// TIA Portal V21 export
// export: Created 2026-11-03T19:44:49.0635428Z, ExportSetting WithDefaults, WithReadOnly, DisplayName Totally Integrated Automation Portal, DisplayVersion V21, DisplayName STEP 7 Professional, DisplayVersion V21, DisplayName STEP 7 Safety, DisplayVersion V21, DisplayName Tech WebApplication, DisplayVersion V21, DisplayName WinCC Basic/Comfort/Advanced, DisplayVersion V21, DisplayName WinCC Professional, DisplayVersion V21, DisplayName WinCC Unified, DisplayVersion V21
DATA_BLOCK "DB_FAT_Demo"   // DB1
{ S7_Optimized_Access := 'FALSE' }
VERSION : 1.0
// SPDX-License-Identifier: MIT. Public passive laboratory example.
// stored: AutoNumber true, CodeModifiedDate 2026-11-03T19:44:32.7091278Z, CompileDate 2026-11-03T19:44:33.4739621Z, CreationDate 2026-11-03T19:44:31.2051572Z, DBAccessibleFromOPCUA true, DBAccessibleFromWebserver true, DownloadDate 0001-01-01T00:00:00Z, InterfaceModifiedDate 2026-11-03T19:44:32.7091278Z, IsConsistent true, IsKnowHowProtected false, IsOnlyStoredInLoadMemory false, IsPLCDB false, IsWriteProtectedInAS false, LoadMemoryLength 5286, ModifiedDate 2026-11-03T19:44:32.7091278Z, ParameterModified 2026-11-03T19:44:32.7091278Z, StructureModified 2026-11-03T19:44:32.7091278Z, WorkMemoryLength 192
   VAR RETAIN
      EnableDemo { ExternalAccessible := 'False'; ExternalVisible := 'False'; ExternalWritable := 'False'} : Bool := TRUE;   // isolated virtual copy only
      StopHealthy : Bool := TRUE;
      P101_Request : Bool := FALSE;
      P101_RequestedSpeed : Real := REAL#60.0;
      P101_RunCommand { ExternalWritable := 'False'} : Bool := FALSE;
      P101_SpeedCommand { ExternalWritable := 'False'} : Real := REAL#0.0;
      P101_Running : Bool := FALSE;
      P101_SpeedFeedback : Real := REAL#0.0;
      P101_Fault : Bool := FALSE;
      P201_Request : Bool := FALSE;
      P201_RequestedSpeed : Real := REAL#60.0;
      P201_RunCommand { ExternalWritable := 'False'} : Bool := FALSE;
      P201_SpeedCommand { ExternalWritable := 'False'} : Real := REAL#0.0;
      P201_Running : Bool := FALSE;
      P201_SpeedFeedback : Real := REAL#0.0;
      P201_Fault : Bool := FALSE;
      P202_Request : Bool := FALSE;
      P202_RequestedSpeed : Real := REAL#60.0;
      P202_RunCommand { ExternalWritable := 'False'} : Bool := FALSE;
      P202_SpeedCommand { ExternalWritable := 'False'} : Real := REAL#0.0;
      P202_Running : Bool := FALSE;
      P202_SpeedFeedback : Real := REAL#0.0;
      P202_Fault : Bool := FALSE;
      P301_Request : Bool := FALSE;
      P301_RequestedSpeed : Real := REAL#60.0;
      P301_RunCommand { ExternalWritable := 'False'} : Bool := FALSE;
      P301_SpeedCommand { ExternalWritable := 'False'} : Real := REAL#0.0;
      P301_Running : Bool := FALSE;
      P301_SpeedFeedback : Real := REAL#0.0;
      P301_Fault : Bool := FALSE;
      XV101_Request : Bool := FALSE;
      XV101_OpenCommand { ExternalWritable := 'False'} : Bool := FALSE;
      XV101_Open : Bool := FALSE;
      XV101_Closed : Bool := TRUE;
      XV201_Request : Bool := FALSE;
      XV201_OpenCommand { ExternalWritable := 'False'} : Bool := FALSE;
      XV201_Open : Bool := FALSE;
      XV201_Closed : Bool := TRUE;
      XV202_Request : Bool := FALSE;
      XV202_OpenCommand { ExternalWritable := 'False'} : Bool := FALSE;
      XV202_Open : Bool := FALSE;
      XV202_Closed : Bool := TRUE;
      XV301_Request : Bool := FALSE;
      XV301_OpenCommand { ExternalWritable := 'False'} : Bool := FALSE;
      XV301_Open : Bool := FALSE;
      XV301_Closed : Bool := TRUE;
      XV102_Request : Bool := FALSE;
      XV102_OpenCommand { ExternalWritable := 'False'} : Bool := FALSE;
      XV102_Open : Bool := FALSE;
      XV102_Closed : Bool := TRUE;
      XV203_Request : Bool := FALSE;
      XV203_OpenCommand { ExternalWritable := 'False'} : Bool := FALSE;
      XV203_Open : Bool := FALSE;
      XV203_Closed : Bool := TRUE;
      XV103_Request : Bool := FALSE;
      XV103_OpenCommand { ExternalWritable := 'False'} : Bool := FALSE;
      XV103_Open : Bool := FALSE;
      XV103_Closed : Bool := TRUE;
      FCV302_RequestedPosition : Real := REAL#0.0;
      FCV302_PositionCommand { ExternalWritable := 'False'} : Real := REAL#0.0;
      FCV302_PositionFeedback : Real := REAL#0.0;
      LT101_Raw : Int := INT#16589;
      LT101_Percent { ExternalWritable := 'False'} : Real := REAL#0.0;
      TK101_Volume : Real := REAL#720.0;
      LSL101 : Bool := FALSE;
      LSH101 : Bool := FALSE;
      LT201_Raw : Int := INT#6912;
      LT201_Percent { ExternalWritable := 'False'} : Real := REAL#0.0;
      TK201_Volume : Real := REAL#450.0;
      LSL201 : Bool := FALSE;
      LSH201 : Bool := FALSE;
      LT301_Raw : Int := INT#4147;
      LT301_Percent { ExternalWritable := 'False'} : Real := REAL#0.0;
      TK301_Volume : Real := REAL#180.0;
      LSL301 : Bool := FALSE;
      LSH301 : Bool := FALSE;
   END_VAR
BEGIN
END_DATA_BLOCK
